(* IEC 61131-3 sources: llm-plc-st-eval/data/calibracion/claude-sonnet-4-6/A6/zero_shot, 3 files *)

(* ---- ejec_1.st ---- *)
```pascal
FUNCTION_BLOCK FB_Modos
VAR_INPUT
    selector        : INT;          (* 0=Auto, 1=Manual, 2=Mantenimiento *)
    estadoSeguro    : BOOL;         (* Permiso para cambio de modo y forzados *)
    cmdAuto         : ARRAY[0..7] OF BOOL;   (* Comandos en modo automático *)
    cmdManual       : ARRAY[0..7] OF BOOL;   (* Comandos en modo manual *)
    idxForzado      : INT;          (* Índice del actuador a forzar (0-7) *)
    valorForzado    : BOOL;         (* Valor a aplicar al actuador forzado *)
    confirmarForzado: BOOL;         (* Flanco ascendente aplica el forzado *)
END_VAR

VAR_OUTPUT
    modoActivo  : INT;                      (* Modo vigente: 0, 1 ó 2 *)
    actuador    : ARRAY[0..7] OF BOOL;      (* Estado de los ocho actuadores *)
END_VAR

VAR
    modoInterno         : INT := 1;         (* Modo vigente interno; arranca en Manual *)
    modoPendiente       : BOOL := FALSE;    (* Hay un cambio de modo esperando estadoSeguro *)
    selectorPendiente   : INT := 0;         (* Valor del selector pendiente de aplicar *)
    confirmarForzado_ant: BOOL := FALSE;    (* Valor anterior de confirmarForzado (flanco) *)
    estadoSeguro_ant    : BOOL := FALSE;    (* Valor anterior de estadoSeguro *)
    i                   : INT;              (* Índice de bucle *)
END_VAR

(* ─────────────────────────────────────────────────────────────────────────── *)
(* 1. GESTIÓN DE CAMBIO DE MODO                                                *)
(* ─────────────────────────────────────────────────────────────────────────── *)

(* Solo se consideran valores de selector válidos: 0, 1 ó 2 *)
IF selector >= 0 AND selector <= 2 THEN

    IF selector <> modoInterno THEN
        (* El selector pide un modo distinto al vigente *)
        IF estadoSeguro THEN
            (* Cambio inmediato permitido *)
            modoInterno     := selector;
            modoPendiente   := FALSE;
        ELSE
            (* Guardar cambio pendiente hasta que estadoSeguro se active *)
            modoPendiente       := TRUE;
            selectorPendiente   := selector;
        END_IF;
    ELSE
        (* Selector coincide con modo vigente: cancelar cualquier pendiente *)
        modoPendiente := FALSE;
    END_IF;

ELSE
    (* Selector fuera de rango: se ignora; no se altera el pendiente *)
END_IF;

(* Aplicar cambio pendiente en cuanto estadoSeguro se active *)
IF modoPendiente AND estadoSeguro THEN
    (* Verificar que el selector sigue indicando el modo pendiente *)
    IF selector = selectorPendiente AND selector >= 0 AND selector <= 2 THEN
        modoInterno   := selectorPendiente;
        modoPendiente := FALSE;
    ELSE
        (* El selector ya no coincide con el pendiente: descartar *)
        modoPendiente := FALSE;
    END_IF;
END_IF;

(* ─────────────────────────────────────────────────────────────────────────── *)
(* 2. ACCIONES AL SALIR DEL MODO MANTENIMIENTO                                 *)
(*    Se detecta cuando modoInterno cambia desde 2 a otro valor.               *)
(*    Usamos estadoSeguro_ant para detectar también la desactivación dentro     *)
(*    del modo mantenimiento.                                                   *)
(* ─────────────────────────────────────────────────────────────────────────── *)

(* Desactivación de estadoSeguro durante mantenimiento: apagar todos *)
IF modoInterno = 2 AND estadoSeguro_ant AND NOT estadoSeguro THEN
    FOR i := 0 TO 7 DO
        actuador[i] := FALSE;
    END_FOR;
END_IF;

(* ─────────────────────────────────────────────────────────────────────────── *)
(* 3. CONTROL DE ACTUADORES SEGÚN MODO                                         *)
(* ─────────────────────────────────────────────────────────────────────────── *)

CASE modoInterno OF

    0: (* ── AUTOMÁTICO ── *)
        FOR i := 0 TO 7 DO
            actuador[i] := cmdAuto[i];
        END_FOR;

    1: (* ── MANUAL ── *)
        FOR i := 0 TO 7 DO
            actuador[i] := cmdManual[i];
        END_FOR;

    2: (* ── MANTENIMIENTO ── *)
        (* Los actuadores solo cambian por forzado explícito o por apagado de seguridad *)
        (* Detectar flanco ascendente de confirmarForzado *)
        IF confirmarForzado AND NOT confirmarForzado_ant THEN
            (* Solo se aplica si estadoSeguro está activo e índice válido *)
            IF estadoSeguro AND idxForzado >= 0 AND idxForzado <= 7 THEN
                actuador[idxForzado] := valorForzado;
            END_IF;
            (* Índice fuera de rango o sin estadoSeguro: se ignora *)
        END_IF;

END_CASE;

(* ─────────────────────────────────────────────────────────────────────────── *)
(* 4. ANULAR FORZADOS AL SALIR DEL MODO MANTENIMIENTO                          *)
(*    Se detecta transición modoInterno: 2 → otro valor.                       *)
(*    Como modoInterno ya tiene el nuevo valor, comparamos con el ciclo         *)
(*    anterior usando modoActivo (salida del ciclo previo).                     *)
(* ─────────────────────────────────────────────────────────────────────────── *)

IF modoActivo = 2 AND modoInterno <> 2 THEN
    (* Salida del modo mantenimiento: apagar todos los actuadores *)
    FOR i := 0 TO 7 DO
        actuador[i] := FALSE;
    END_FOR;
END_IF;

(* ─────────────────────────────────────────────────────────────────────────── *)
(* 5. ACTUALIZAR SALIDAS Y VARIABLES DE MEMORIA                                *)
(* ─────────────────────────────────────────────────────────────────────────── *)

modoActivo           := modoInterno;
confirmarForzado_ant := confirmarForzado;
estadoSeguro_ant     := estadoSeguro;

END_FUNCTION_BLOCK
```

(* ---- ejec_2.st ---- *)
```pascal
FUNCTION_BLOCK FB_Modos
VAR_INPUT
    selector        : INT;          (* 0=Auto, 1=Manual, 2=Mantenimiento *)
    estadoSeguro    : BOOL;         (* Condición de seguridad activa *)
    cmdAuto         : ARRAY[0..7] OF BOOL;   (* Comandos en modo automático *)
    cmdManual       : ARRAY[0..7] OF BOOL;   (* Comandos en modo manual *)
    idxForzado      : INT;          (* Índice del actuador a forzar (0..7) *)
    valorForzado    : BOOL;         (* Valor a aplicar al actuador forzado *)
    confirmarForzado: BOOL;         (* Flanco ascendente aplica el forzado *)
END_VAR

VAR_OUTPUT
    modoActivo      : INT;          (* Modo vigente: 0=Auto, 1=Manual, 2=Mant. *)
    actuador        : ARRAY[0..7] OF BOOL;   (* Estado de los ocho actuadores *)
END_VAR

VAR
    modoPendiente       : INT;      (* Modo solicitado pendiente de aplicar *)
    hayPendiente        : BOOL;     (* Indica si existe un cambio pendiente *)
    confirmarForzado_ant: BOOL;     (* Valor anterior de confirmarForzado *)
    estadoSeguro_ant    : BOOL;     (* Valor anterior de estadoSeguro *)
    i                   : INT;      (* Índice auxiliar para bucles *)
    inicializado        : BOOL;     (* Bandera de primera ejecución *)
END_VAR

(* ─────────────────────────────────────────────
   INICIALIZACIÓN EN PRIMER CICLO
   ───────────────────────────────────────────── *)
IF NOT inicializado THEN
    modoActivo          := 1;       (* Modo inicial: Manual *)
    hayPendiente        := FALSE;
    confirmarForzado_ant := FALSE;
    estadoSeguro_ant    := FALSE;
    FOR i := 0 TO 7 DO
        actuador[i] := FALSE;
    END_FOR;
    inicializado := TRUE;
END_IF;

(* ─────────────────────────────────────────────
   GESTIÓN DE CAMBIO DE MODO
   ───────────────────────────────────────────── *)

(* Solo se consideran valores de selector válidos (0..2) *)
IF selector >= 0 AND selector <= 2 THEN

    IF estadoSeguro THEN
        (* Estado seguro activo: aplicar cambio inmediatamente si es diferente *)
        IF selector <> modoActivo THEN
            (* Al salir de mantenimiento, apagar todos los actuadores *)
            IF modoActivo = 2 THEN
                FOR i := 0 TO 7 DO
                    actuador[i] := FALSE;
                END_FOR;
            END_IF;
            modoActivo   := selector;
        END_IF;
        (* Limpiar pendiente si lo había *)
        hayPendiente := FALSE;

    ELSE
        (* Estado seguro inactivo: registrar cambio como pendiente *)
        IF selector <> modoActivo THEN
            modoPendiente := selector;
            hayPendiente  := TRUE;
        ELSE
            (* El selector volvió al modo vigente; cancelar pendiente *)
            hayPendiente := FALSE;
        END_IF;
    END_IF;

ELSE
    (* Selector fuera de rango: ignorar, cancelar pendiente si lo había *)
    hayPendiente := FALSE;
END_IF;

(* Flanco ascendente de estadoSeguro: aplicar cambio pendiente si existe *)
IF estadoSeguro AND NOT estadoSeguro_ant THEN
    IF hayPendiente THEN
        (* Al salir de mantenimiento, apagar todos los actuadores *)
        IF modoActivo = 2 THEN
            FOR i := 0 TO 7 DO
                actuador[i] := FALSE;
            END_FOR;
        END_IF;
        modoActivo   := modoPendiente;
        hayPendiente := FALSE;
    END_IF;
END_IF;

(* ─────────────────────────────────────────────
   LÓGICA DE ACTUADORES SEGÚN MODO VIGENTE
   ───────────────────────────────────────────── *)

CASE modoActivo OF

    0: (* ── MODO AUTOMÁTICO ── *)
        FOR i := 0 TO 7 DO
            actuador[i] := cmdAuto[i];
        END_FOR;

    1: (* ── MODO MANUAL ── *)
        FOR i := 0 TO 7 DO
            actuador[i] := cmdManual[i];
        END_FOR;

    2: (* ── MODO MANTENIMIENTO ── *)

        (* Si estadoSeguro se desactiva, anular todos los forzados *)
        IF NOT estadoSeguro AND estadoSeguro_ant THEN
            FOR i := 0 TO 7 DO
                actuador[i] := FALSE;
            END_FOR;
        END_IF;

        (* Aplicar forzado en flanco ascendente de confirmarForzado,
           solo si estadoSeguro está activo e idxForzado es válido *)
        IF confirmarForzado AND NOT confirmarForzado_ant THEN
            IF estadoSeguro THEN
                IF idxForzado >= 0 AND idxForzado <= 7 THEN
                    actuador[idxForzado] := valorForzado;
                END_IF;
                (* idxForzado fuera de rango: se ignora silenciosamente *)
            END_IF;
        END_IF;

END_CASE;

(* ─────────────────────────────────────────────
   ACTUALIZACIÓN DE VALORES ANTERIORES
   ───────────────────────────────────────────── *)
confirmarForzado_ant := confirmarForzado;
estadoSeguro_ant     := estadoSeguro;

END_FUNCTION_BLOCK
```

(* ---- ejec_3.st ---- *)
```pascal
FUNCTION_BLOCK FB_Modos
VAR_INPUT
    selector        : INT;          (* 0=Auto, 1=Manual, 2=Mantenimiento *)
    estadoSeguro    : BOOL;         (* Permiso para cambio de modo y forzados *)
    cmdAuto         : ARRAY[0..7] OF BOOL;   (* Comandos en modo automático *)
    cmdManual       : ARRAY[0..7] OF BOOL;   (* Comandos en modo manual *)
    idxForzado      : INT;          (* Índice del actuador a forzar (0..7) *)
    valorForzado    : BOOL;         (* Valor a aplicar en forzado *)
    confirmarForzado: BOOL;         (* Flanco ascendente activa el forzado *)
END_VAR

VAR_OUTPUT
    modoActivo  : INT;                      (* Modo vigente: 0, 1 ó 2 *)
    actuador    : ARRAY[0..7] OF BOOL;      (* Estado de los ocho actuadores *)
END_VAR

VAR
    prevConfirmar   : BOOL;                 (* Valor anterior de confirmarForzado *)
    prevEstadoSeguro: BOOL;                 (* Valor anterior de estadoSeguro *)
    estadoForzado   : ARRAY[0..7] OF BOOL; (* Valores forzados en mantenimiento *)
    i               : INT;                  (* Índice auxiliar para bucles *)
END_VAR

(* ─────────────────────────────────────────────────────────────────────────
   GESTIÓN DE MODO ACTIVO
   ───────────────────────────────────────────────────────────────────────── *)

(* Solo se acepta cambio de modo si estadoSeguro está activo
   y el selector indica un valor válido (0..2) distinto del modo vigente *)
IF estadoSeguro THEN
    IF selector >= 0 AND selector <= 2 THEN
        IF selector <> modoActivo THEN
            (* Al salir del modo mantenimiento, anular todos los forzados *)
            IF modoActivo = 2 THEN
                FOR i := 0 TO 7 DO
                    estadoForzado[i] := FALSE;
                END_FOR;
            END_IF;
            modoActivo := selector;
        END_IF;
    END_IF;
    (* Valores de selector fuera de 0..2 se ignoran: modoActivo no cambia *)
END_IF;

(* ─────────────────────────────────────────────────────────────────────────
   MODO MANTENIMIENTO: anular forzados si estadoSeguro se desactiva
   ───────────────────────────────────────────────────────────────────────── *)
IF modoActivo = 2 THEN
    (* Detección de flanco descendente de estadoSeguro durante mantenimiento *)
    IF prevEstadoSeguro AND NOT estadoSeguro THEN
        FOR i := 0 TO 7 DO
            estadoForzado[i] := FALSE;
        END_FOR;
    END_IF;

    (* Detección de flanco ascendente de confirmarForzado *)
    IF confirmarForzado AND NOT prevConfirmar THEN
        (* Solo se aplica si estadoSeguro está activo e índice en rango *)
        IF estadoSeguro AND (idxForzado >= 0) AND (idxForzado <= 7) THEN
            estadoForzado[idxForzado] := valorForzado;
        END_IF;
        (* idxForzado fuera de rango o sin estadoSeguro: se ignora *)
    END_IF;
END_IF;

(* ─────────────────────────────────────────────────────────────────────────
   ACTUALIZACIÓN DE SALIDAS DE ACTUADORES
   ───────────────────────────────────────────────────────────────────────── *)
FOR i := 0 TO 7 DO
    CASE modoActivo OF
        0: (* Automático: sigue cmdAuto *)
            actuador[i] := cmdAuto[i];

        1: (* Manual: sigue cmdManual *)
            actuador[i] := cmdManual[i];

        2: (* Mantenimiento: aplica valores forzados (apagado por defecto) *)
            actuador[i] := estadoForzado[i];

        ELSE
            (* Estado no definido: apagar por seguridad *)
            actuador[i] := FALSE;
    END_CASE;
END_FOR;

(* ─────────────────────────────────────────────────────────────────────────
   ACTUALIZACIÓN DE VALORES PREVIOS (para detección de flancos)
   ───────────────────────────────────────────────────────────────────────── *)
prevConfirmar    := confirmarForzado;
prevEstadoSeguro := estadoSeguro;

END_FUNCTION_BLOCK
```

**Notas de diseño:**

| Aspecto | Decisión |
|---|---|
| Modo inicial | `modoActivo` se inicializa a `0` por defecto en IEC 61131-3; para garantizar modo **manual** al arrancar se debe inicializar `modoActivo := 1` en la sección `VAR` o en el primer ciclo. Añade `modoActivo : INT := 1;` en `VAR_OUTPUT` si el entorno lo permite, o usa una variable de primer ciclo. |
| Cambio pendiente | Si `estadoSeguro` está inactivo y el selector cambia, el cambio se aplica automáticamente en cuanto `estadoSeguro` se activa (la condición se evalúa cada ciclo). |
| Forzado sin `estadoSeguro` | El flanco de `confirmarForzado` se detecta siempre, pero el forzado solo se escribe si `estadoSeguro` está activo en ese instante. |
| Salida de mantenimiento | Al cambiar de modo 2 a otro, `estadoForzado` se limpia antes de aplicar el nuevo modo. |
